TYPE "ST_SequenceAnnotation"
VERSION : 0.1
   STRUCT
      "RowIdx" : Int;
      "IsError" : Bool;
      "Key" : String[120];
      "SourcePath" : String[80];
   END_STRUCT;
END_TYPE
